// Mitsubishi GX Works2 project: plc_v1   PLC: Q03UDV

PROGRAM COM_RACK
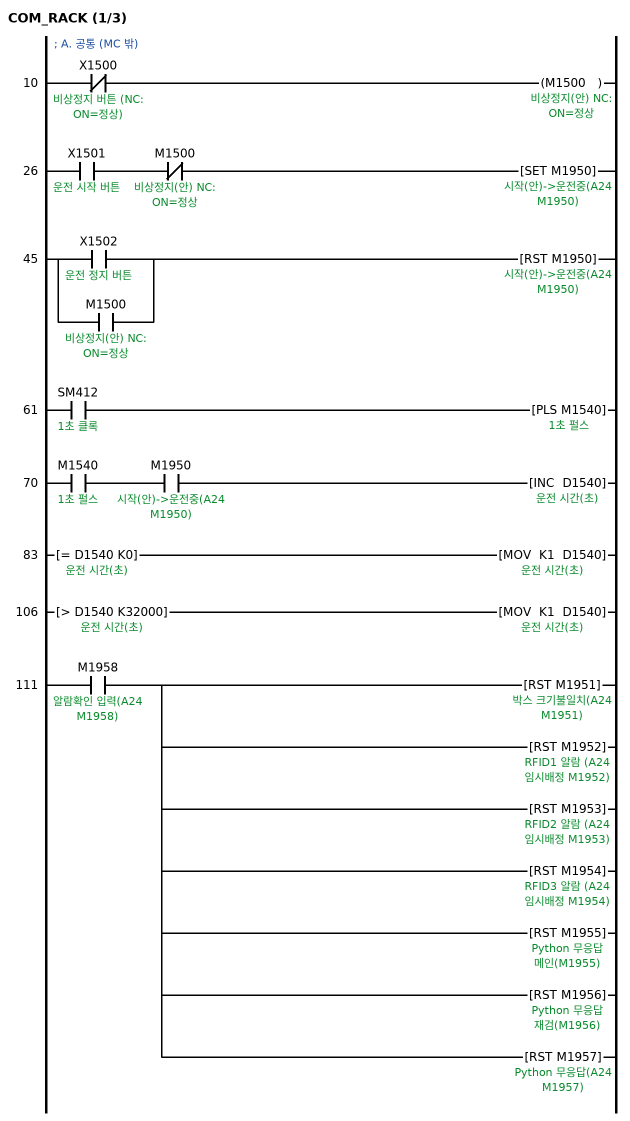
; A. 공통 (MC 밖)
10    LDI     X1500  ; 비상정지 버튼 (NC: ON=정상)
      OUT     M1500  ; 비상정지(안) NC: ON=정상
        [note] 비상정지(안) NC: ON=정상
26    LD      X1501  ; 운전 시작 버튼
      ANI     M1500  ; 비상정지(안) NC: ON=정상
      SET     M1950  ; 시작(안)->운전중(A24 M1950)
        [note] 시작(안)->운전중(A24 M1950)
45    LD      X1502  ; 운전 정지 버튼
      OR      M1500  ; 비상정지(안) NC: ON=정상
      RST     M1950  ; 시작(안)->운전중(A24 M1950)
        [note] 정지(안) 또는 비상정지
61    LD      SM412  ; 1초 클록
      PLS     M1540  ; 1초 펄스
        [note] 1초 펄스
70    LD      M1540  ; 1초 펄스
      AND     M1950  ; 시작(안)->운전중(A24 M1950)
      INC     D1540  ; 운전 시간(초)
        [note] 운전 시간(초)
83    LD=     D1540 K0  ; 운전 시간(초)
      MOV     K1 D1540
        [note] 0은 입고 중 표시로 쓰므로 1부터
106   LD>     D1540 K32000  ; 운전 시간(초)
      MOV     K1 D1540
111   LD      M1958  ; 알람확인 입력(A24 M1958)
      RST     M1951  ; 박스 크기불일치(A24 M1951)
      RST     M1952  ; RFID1 알람 (A24 임시배정 M1952)
      RST     M1953  ; RFID2 알람 (A24 임시배정 M1953)
      RST     M1954  ; RFID3 알람 (A24 임시배정 M1954)
      RST     M1955  ; Python 무응답 메인(M1955)
      RST     M1956  ; Python 무응답 재검(M1956)
      RST     M1957  ; Python 무응답(A24 M1957)
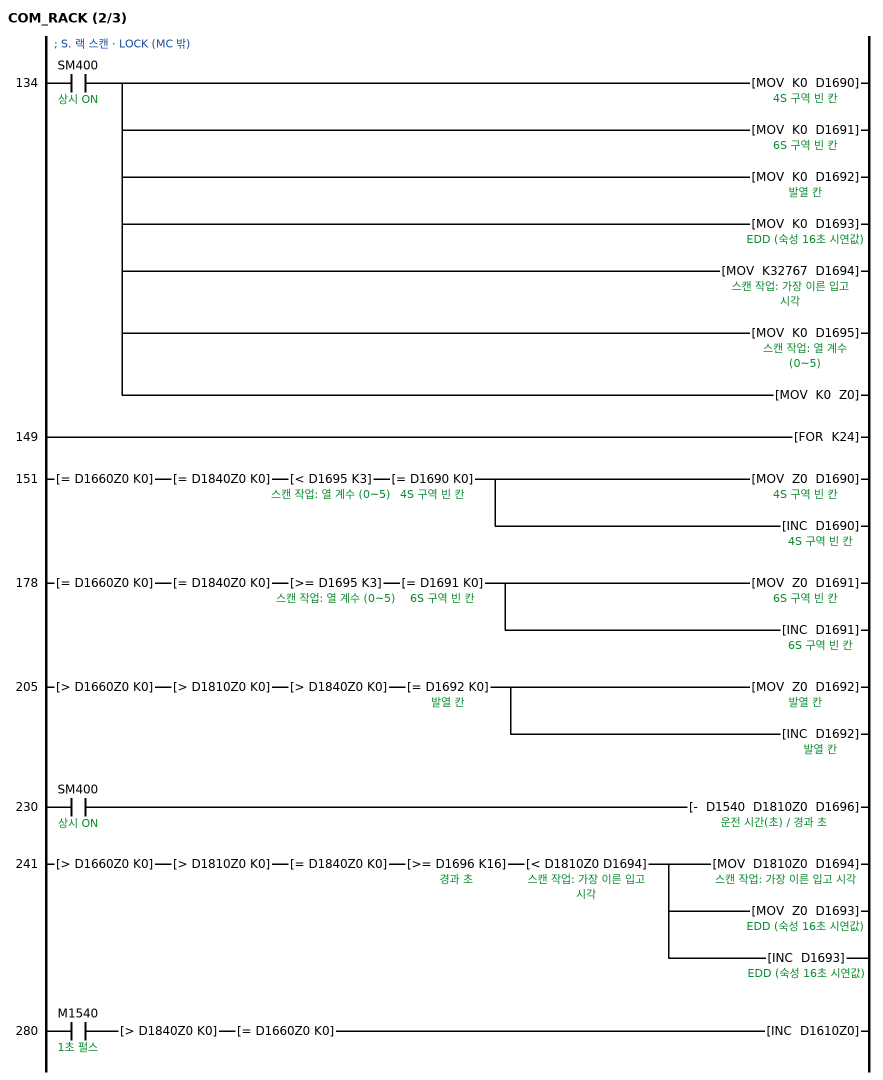
; S. 랙 스캔 · LOCK (MC 밖)
134   LD      SM400  ; 상시 ON
      MOV     K0 D1690  ; 4S 구역 빈 칸
      MOV     K0 D1691  ; 6S 구역 빈 칸
      MOV     K0 D1692  ; 발열 칸
      MOV     K0 D1693  ; EDD (숙성 16초 시연값)
      MOV     K32767 D1694  ; 스캔 작업: 가장 이른 입고 시각
      MOV     K0 D1695  ; 스캔 작업: 열 계수 (0~5)
      MOV     K0 Z0
149   FOR     K24
151   LD=     D1660Z0 K0
      AND=    D1840Z0 K0
      AND<    D1695 K3  ; 스캔 작업: 열 계수 (0~5)
      AND=    D1690 K0  ; 4S 구역 빈 칸
      MOV     Z0 D1690
      INC     D1690
        [note] 4S 구역 빈 칸
178   LD=     D1660Z0 K0
      AND=    D1840Z0 K0
      AND>=   D1695 K3  ; 스캔 작업: 열 계수 (0~5)
      AND=    D1691 K0  ; 6S 구역 빈 칸
      MOV     Z0 D1691
      INC     D1691
        [note] 6S 구역 빈 칸
205   LD>     D1660Z0 K0
      AND>    D1810Z0 K0
      AND>    D1840Z0 K0
      AND=    D1692 K0  ; 발열 칸
      MOV     Z0 D1692
      INC     D1692
        [note] 발열 칸
230   LD      SM400  ; 상시 ON
      -       D1540 D1810Z0 D1696  ; 경과 초
        [note] 경과 초
241   LD>     D1660Z0 K0
      AND>    D1810Z0 K0
      AND=    D1840Z0 K0
      AND>=   D1696 K16  ; 경과 초
      AND<    D1810Z0 D1694  ; 스캔 작업: 가장 이른 입고 시각
      MOV     D1810Z0 D1694
      MOV     Z0 D1693
      INC     D1693
        [note] EDD (숙성 16초 시연값)
280   LD      M1540  ; 1초 펄스
      AND>    D1840Z0 K0
      AND=    D1660Z0 K0
      INC     D1610Z0
        [note] LOCK 경과(초)
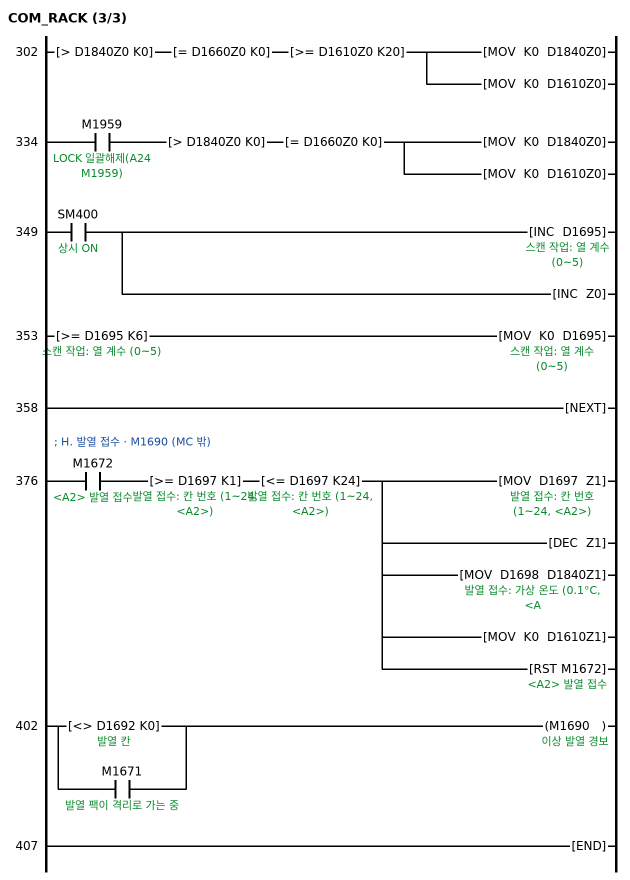
302   LD>     D1840Z0 K0
      AND=    D1660Z0 K0
      AND>=   D1610Z0 K20
      MOV     K0 D1840Z0
      MOV     K0 D1610Z0
        [note] 20초 뒤 자동 해제 (D13)
334   LD      M1959  ; LOCK 일괄해제(A24 M1959)
      AND>    D1840Z0 K0
      AND=    D1660Z0 K0
      MOV     K0 D1840Z0
      MOV     K0 D1610Z0
349   LD      SM400  ; 상시 ON
      INC     D1695
      INC     Z0
353   LD>=    D1695 K6  ; 스캔 작업: 열 계수 (0~5)
      MOV     K0 D1695
358   NEXT
; H. 발열 접수 · M1690 (MC 밖)
376   LD      M1672  ; <A2> 발열 접수
      AND>=   D1697 K1  ; 발열 접수: 칸 번호 (1~24, <A2>)
      AND<=   D1697 K24  ; 발열 접수: 칸 번호 (1~24, <A2>)
      MOV     D1697 Z1
      DEC     Z1
      MOV     D1698 D1840Z1  ; 발열 접수: 가상 온도 (0.1°C, <A
      MOV     K0 D1610Z1
      RST     M1672  ; <A2> 발열 접수
        [note] <A2> 발열 접수
402   LD<>    D1692 K0  ; 발열 칸
      OR      M1671  ; 발열 팩이 격리로 가는 중
      OUT     M1690  ; 이상 발열 경보
407   END
END_PROGRAM

PROGRAM MC_MAIN
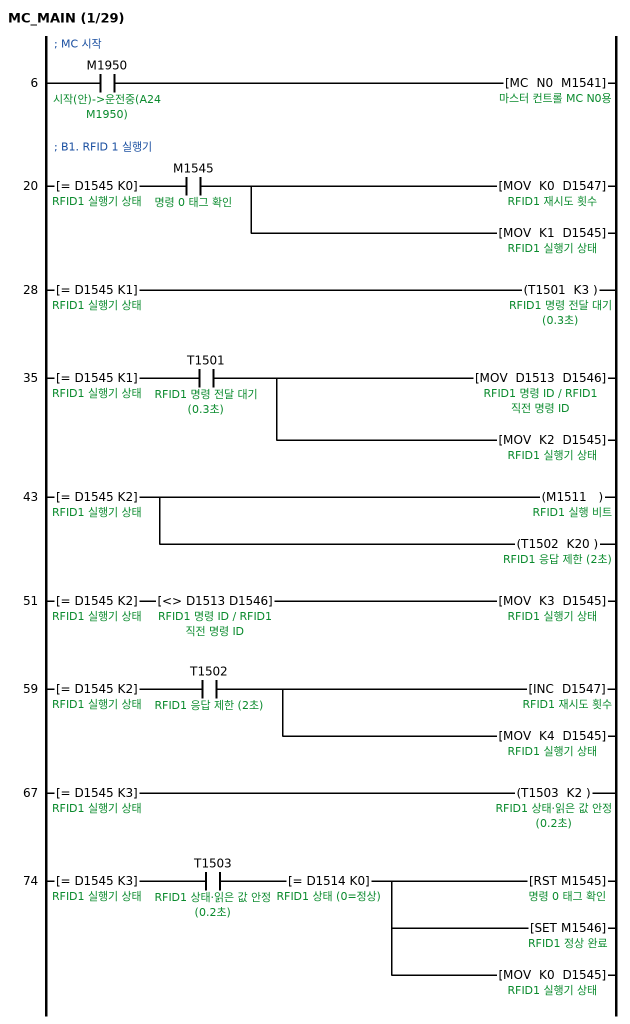
; MC 시작
6     LD      M1950  ; 시작(안)->운전중(A24 M1950)
      MC      N0 M1541  ; 마스터 컨트롤 MC N0용
; B1. RFID 1 실행기
20    LD=     D1545 K0  ; RFID1 실행기 상태
      AND     M1545  ; 명령 0 태그 확인
      MOV     K0 D1547  ; RFID1 재시도 횟수
      MOV     K1 D1545
28    LD=     D1545 K1  ; RFID1 실행기 상태
      OUT     T1501 K3  ; RFID1 명령 전달 대기 (0.3초)
35    LD=     D1545 K1  ; RFID1 실행기 상태
      AND     T1501  ; RFID1 명령 전달 대기 (0.3초)
      MOV     D1513 D1546  ; RFID1 명령 ID / RFID1 직전 명령 ID
      MOV     K2 D1545
43    LD=     D1545 K2  ; RFID1 실행기 상태
      OUT     M1511  ; RFID1 실행 비트
      OUT     T1502 K20  ; RFID1 응답 제한 (2초)
51    LD=     D1545 K2  ; RFID1 실행기 상태
      AND<>   D1513 D1546  ; RFID1 명령 ID / RFID1 직전 명령 ID
      MOV     K3 D1545
59    LD=     D1545 K2  ; RFID1 실행기 상태
      AND     T1502  ; RFID1 응답 제한 (2초)
      INC     D1547
      MOV     K4 D1545
67    LD=     D1545 K3  ; RFID1 실행기 상태
      OUT     T1503 K2  ; RFID1 상태·읽은 값 안정 (0.2초)
74    LD=     D1545 K3  ; RFID1 실행기 상태
      AND     T1503  ; RFID1 상태·읽은 값 안정 (0.2초)
      AND=    D1514 K0  ; RFID1 상태 (0=정상)
      RST     M1545  ; 명령 0 태그 확인
      SET     M1546  ; RFID1 정상 완료
      MOV     K0 D1545
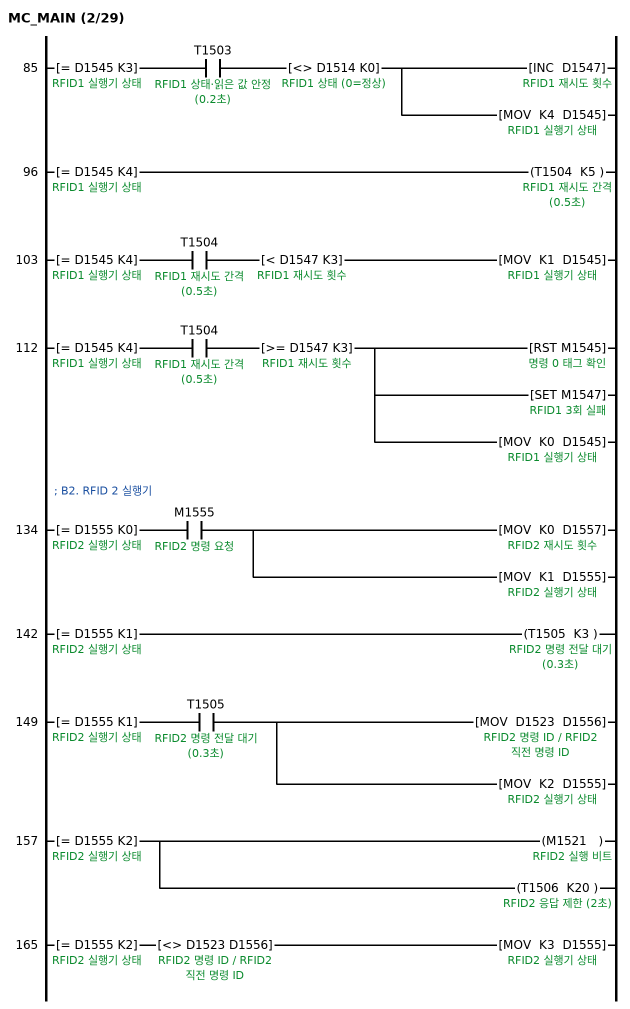
85    LD=     D1545 K3  ; RFID1 실행기 상태
      AND     T1503  ; RFID1 상태·읽은 값 안정 (0.2초)
      AND<>   D1514 K0  ; RFID1 상태 (0=정상)
      INC     D1547
      MOV     K4 D1545
96    LD=     D1545 K4  ; RFID1 실행기 상태
      OUT     T1504 K5  ; RFID1 재시도 간격 (0.5초)
103   LD=     D1545 K4  ; RFID1 실행기 상태
      AND     T1504  ; RFID1 재시도 간격 (0.5초)
      AND<    D1547 K3  ; RFID1 재시도 횟수
      MOV     K1 D1545
112   LD=     D1545 K4  ; RFID1 실행기 상태
      AND     T1504  ; RFID1 재시도 간격 (0.5초)
      AND>=   D1547 K3  ; RFID1 재시도 횟수
      RST     M1545  ; 명령 0 태그 확인
      SET     M1547  ; RFID1 3회 실패
      MOV     K0 D1545
; B2. RFID 2 실행기
134   LD=     D1555 K0  ; RFID2 실행기 상태
      AND     M1555  ; RFID2 명령 요청
      MOV     K0 D1557  ; RFID2 재시도 횟수
      MOV     K1 D1555
142   LD=     D1555 K1  ; RFID2 실행기 상태
      OUT     T1505 K3  ; RFID2 명령 전달 대기 (0.3초)
149   LD=     D1555 K1  ; RFID2 실행기 상태
      AND     T1505  ; RFID2 명령 전달 대기 (0.3초)
      MOV     D1523 D1556  ; RFID2 명령 ID / RFID2 직전 명령 ID
      MOV     K2 D1555
157   LD=     D1555 K2  ; RFID2 실행기 상태
      OUT     M1521  ; RFID2 실행 비트
      OUT     T1506 K20  ; RFID2 응답 제한 (2초)
165   LD=     D1555 K2  ; RFID2 실행기 상태
      AND<>   D1523 D1556  ; RFID2 명령 ID / RFID2 직전 명령 ID
      MOV     K3 D1555
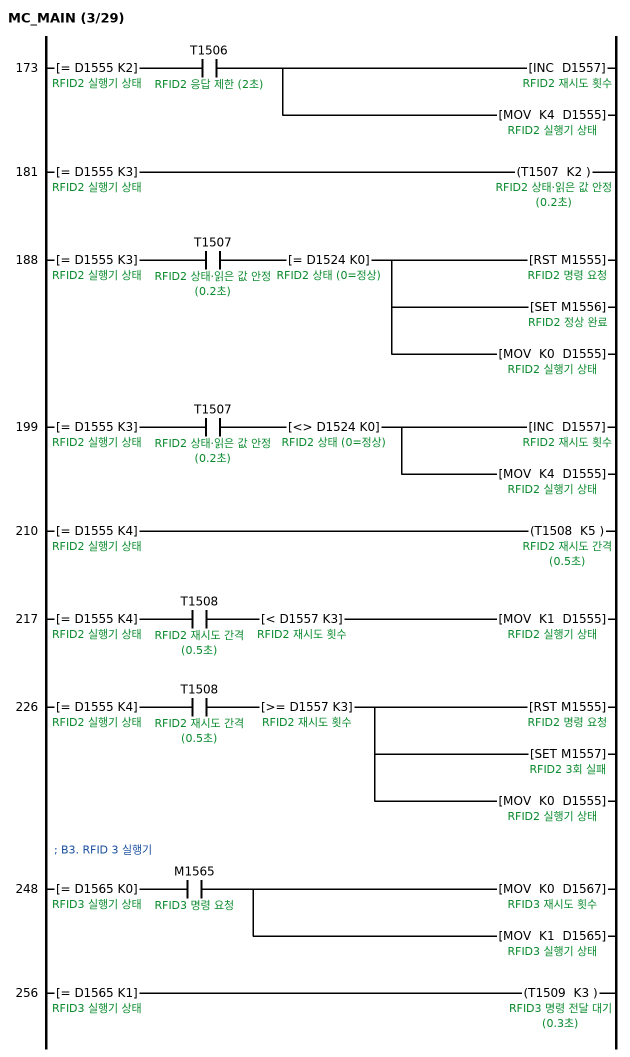
173   LD=     D1555 K2  ; RFID2 실행기 상태
      AND     T1506  ; RFID2 응답 제한 (2초)
      INC     D1557
      MOV     K4 D1555
181   LD=     D1555 K3  ; RFID2 실행기 상태
      OUT     T1507 K2  ; RFID2 상태·읽은 값 안정 (0.2초)
188   LD=     D1555 K3  ; RFID2 실행기 상태
      AND     T1507  ; RFID2 상태·읽은 값 안정 (0.2초)
      AND=    D1524 K0  ; RFID2 상태 (0=정상)
      RST     M1555  ; RFID2 명령 요청
      SET     M1556  ; RFID2 정상 완료
      MOV     K0 D1555
199   LD=     D1555 K3  ; RFID2 실행기 상태
      AND     T1507  ; RFID2 상태·읽은 값 안정 (0.2초)
      AND<>   D1524 K0  ; RFID2 상태 (0=정상)
      INC     D1557
      MOV     K4 D1555
210   LD=     D1555 K4  ; RFID2 실행기 상태
      OUT     T1508 K5  ; RFID2 재시도 간격 (0.5초)
217   LD=     D1555 K4  ; RFID2 실행기 상태
      AND     T1508  ; RFID2 재시도 간격 (0.5초)
      AND<    D1557 K3  ; RFID2 재시도 횟수
      MOV     K1 D1555
226   LD=     D1555 K4  ; RFID2 실행기 상태
      AND     T1508  ; RFID2 재시도 간격 (0.5초)
      AND>=   D1557 K3  ; RFID2 재시도 횟수
      RST     M1555  ; RFID2 명령 요청
      SET     M1557  ; RFID2 3회 실패
      MOV     K0 D1555
; B3. RFID 3 실행기
248   LD=     D1565 K0  ; RFID3 실행기 상태
      AND     M1565  ; RFID3 명령 요청
      MOV     K0 D1567  ; RFID3 재시도 횟수
      MOV     K1 D1565
256   LD=     D1565 K1  ; RFID3 실행기 상태
      OUT     T1509 K3  ; RFID3 명령 전달 대기 (0.3초)
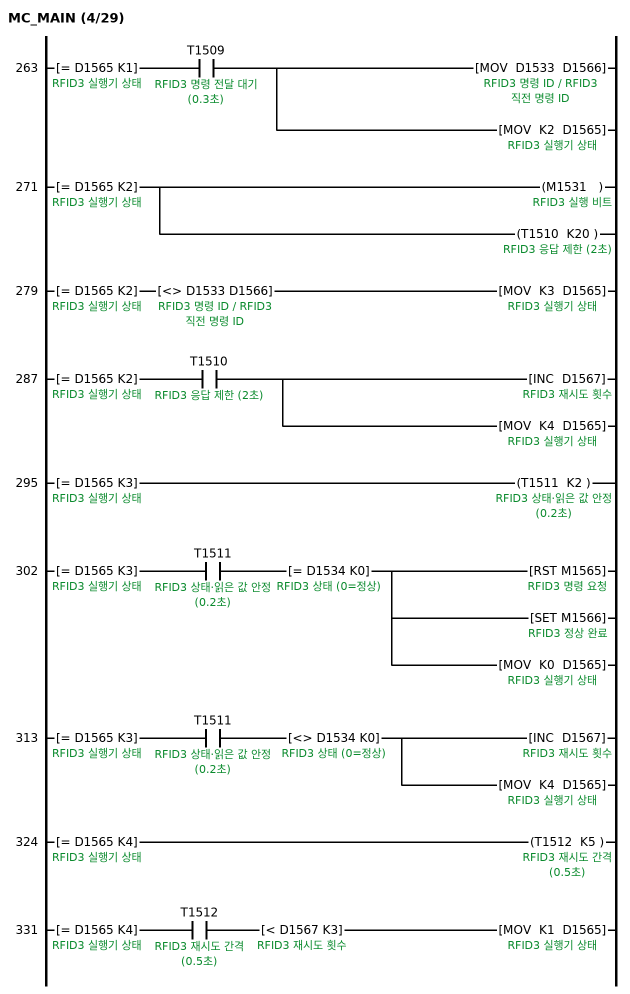
263   LD=     D1565 K1  ; RFID3 실행기 상태
      AND     T1509  ; RFID3 명령 전달 대기 (0.3초)
      MOV     D1533 D1566  ; RFID3 명령 ID / RFID3 직전 명령 ID
      MOV     K2 D1565
271   LD=     D1565 K2  ; RFID3 실행기 상태
      OUT     M1531  ; RFID3 실행 비트
      OUT     T1510 K20  ; RFID3 응답 제한 (2초)
279   LD=     D1565 K2  ; RFID3 실행기 상태
      AND<>   D1533 D1566  ; RFID3 명령 ID / RFID3 직전 명령 ID
      MOV     K3 D1565
287   LD=     D1565 K2  ; RFID3 실행기 상태
      AND     T1510  ; RFID3 응답 제한 (2초)
      INC     D1567
      MOV     K4 D1565
295   LD=     D1565 K3  ; RFID3 실행기 상태
      OUT     T1511 K2  ; RFID3 상태·읽은 값 안정 (0.2초)
302   LD=     D1565 K3  ; RFID3 실행기 상태
      AND     T1511  ; RFID3 상태·읽은 값 안정 (0.2초)
      AND=    D1534 K0  ; RFID3 상태 (0=정상)
      RST     M1565  ; RFID3 명령 요청
      SET     M1566  ; RFID3 정상 완료
      MOV     K0 D1565
313   LD=     D1565 K3  ; RFID3 실행기 상태
      AND     T1511  ; RFID3 상태·읽은 값 안정 (0.2초)
      AND<>   D1534 K0  ; RFID3 상태 (0=정상)
      INC     D1567
      MOV     K4 D1565
324   LD=     D1565 K4  ; RFID3 실행기 상태
      OUT     T1512 K5  ; RFID3 재시도 간격 (0.5초)
331   LD=     D1565 K4  ; RFID3 실행기 상태
      AND     T1512  ; RFID3 재시도 간격 (0.5초)
      AND<    D1567 K3  ; RFID3 재시도 횟수
      MOV     K1 D1565
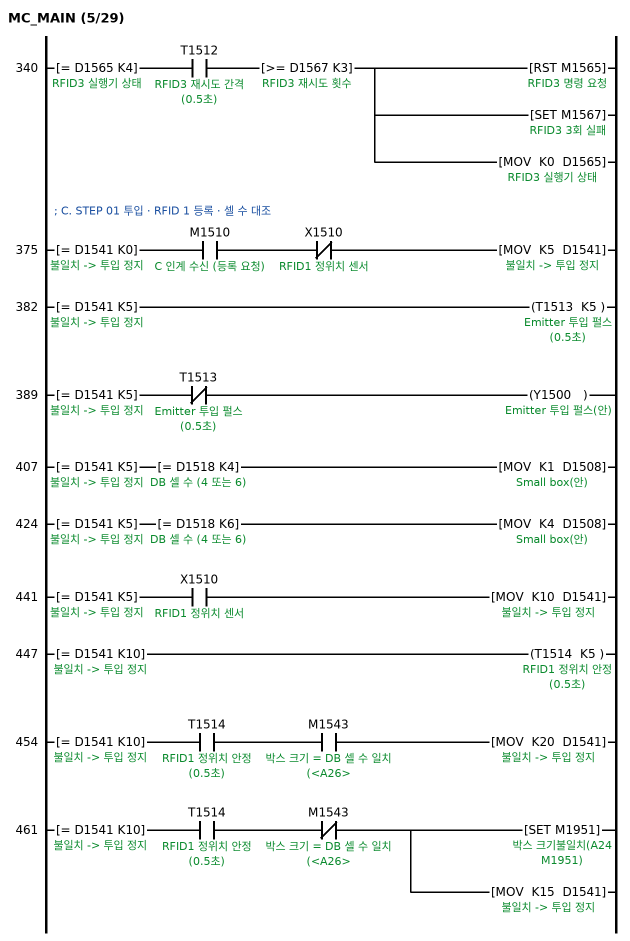
340   LD=     D1565 K4  ; RFID3 실행기 상태
      AND     T1512  ; RFID3 재시도 간격 (0.5초)
      AND>=   D1567 K3  ; RFID3 재시도 횟수
      RST     M1565  ; RFID3 명령 요청
      SET     M1567  ; RFID3 3회 실패
      MOV     K0 D1565
; C. STEP 01 투입 · RFID 1 등록 · 셀 수 대조
375   LD=     D1541 K0  ; 불일치 -> 투입 정지
      AND     M1510  ; C 인계 수신 (등록 요청)
      ANI     X1510  ; RFID1 정위치 센서
      MOV     K5 D1541
382   LD=     D1541 K5  ; 불일치 -> 투입 정지
      OUT     T1513 K5  ; Emitter 투입 펄스 (0.5초)
389   LD=     D1541 K5  ; 불일치 -> 투입 정지
      ANI     T1513  ; Emitter 투입 펄스 (0.5초)
      OUT     Y1500  ; Emitter 투입 펄스(안)
        [note] Emitter 투입 펄스(안)
407   LD=     D1541 K5  ; 불일치 -> 투입 정지
      AND=    D1518 K4  ; DB 셀 수 (4 또는 6)
      MOV     K1 D1508  ; Small box(안)
        [note] Small box(안)
424   LD=     D1541 K5  ; 불일치 -> 투입 정지
      AND=    D1518 K6  ; DB 셀 수 (4 또는 6)
      MOV     K4 D1508
        [note] Large box(안)
441   LD=     D1541 K5  ; 불일치 -> 투입 정지
      AND     X1510  ; RFID1 정위치 센서
      MOV     K10 D1541
447   LD=     D1541 K10  ; 불일치 -> 투입 정지
      OUT     T1514 K5  ; RFID1 정위치 안정 (0.5초)
454   LD=     D1541 K10  ; 불일치 -> 투입 정지
      AND     T1514  ; RFID1 정위치 안정 (0.5초)
      AND     M1543  ; 박스 크기 = DB 셀 수 일치 (<A26>
      MOV     K20 D1541
461   LD=     D1541 K10  ; 불일치 -> 투입 정지
      AND     T1514  ; RFID1 정위치 안정 (0.5초)
      ANI     M1543  ; 박스 크기 = DB 셀 수 일치 (<A26>
      SET     M1951  ; 박스 크기불일치(A24 M1951)
        [note] 박스 크기불일치(A24 M1951)
      MOV     K15 D1541
        [note] 불일치 -> 투입 정지
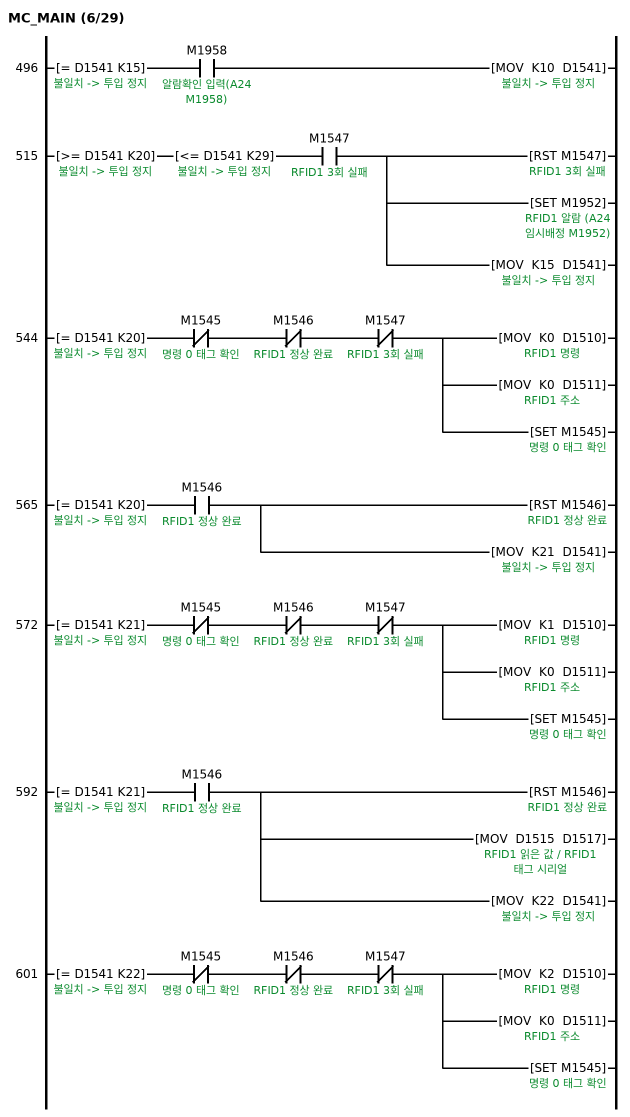
496   LD=     D1541 K15  ; 불일치 -> 투입 정지
      AND     M1958  ; 알람확인 입력(A24 M1958)
      MOV     K10 D1541
        [note] 알람 확인 뒤 다시 대조
515   LD>=    D1541 K20  ; 불일치 -> 투입 정지
      AND<=   D1541 K29  ; 불일치 -> 투입 정지
      AND     M1547  ; RFID1 3회 실패
      RST     M1547  ; RFID1 3회 실패
      SET     M1952  ; RFID1 알람 (A24 임시배정 M1952)
        [note] RFID1 알람 (A24 임시배정 M1952)
      MOV     K15 D1541
544   LD=     D1541 K20  ; 불일치 -> 투입 정지
      ANI     M1545  ; 명령 0 태그 확인
      ANI     M1546  ; RFID1 정상 완료
      ANI     M1547  ; RFID1 3회 실패
      MOV     K0 D1510  ; RFID1 명령
      MOV     K0 D1511  ; RFID1 주소
      SET     M1545  ; 명령 0 태그 확인
        [note] 명령 0 태그 확인
565   LD=     D1541 K20  ; 불일치 -> 투입 정지
      AND     M1546  ; RFID1 정상 완료
      RST     M1546  ; RFID1 정상 완료
      MOV     K21 D1541
572   LD=     D1541 K21  ; 불일치 -> 투입 정지
      ANI     M1545  ; 명령 0 태그 확인
      ANI     M1546  ; RFID1 정상 완료
      ANI     M1547  ; RFID1 3회 실패
      MOV     K1 D1510
      MOV     K0 D1511
      SET     M1545  ; 명령 0 태그 확인
        [note] 명령 1 시리얼
592   LD=     D1541 K21  ; 불일치 -> 투입 정지
      AND     M1546  ; RFID1 정상 완료
      RST     M1546  ; RFID1 정상 완료
      MOV     D1515 D1517  ; RFID1 읽은 값 / RFID1 태그 시리얼
      MOV     K22 D1541
601   LD=     D1541 K22  ; 불일치 -> 투입 정지
      ANI     M1545  ; 명령 0 태그 확인
      ANI     M1546  ; RFID1 정상 완료
      ANI     M1547  ; RFID1 3회 실패
      MOV     K2 D1510
      MOV     K0 D1511
      SET     M1545  ; 명령 0 태그 확인
        [note] 명령 2 idx0
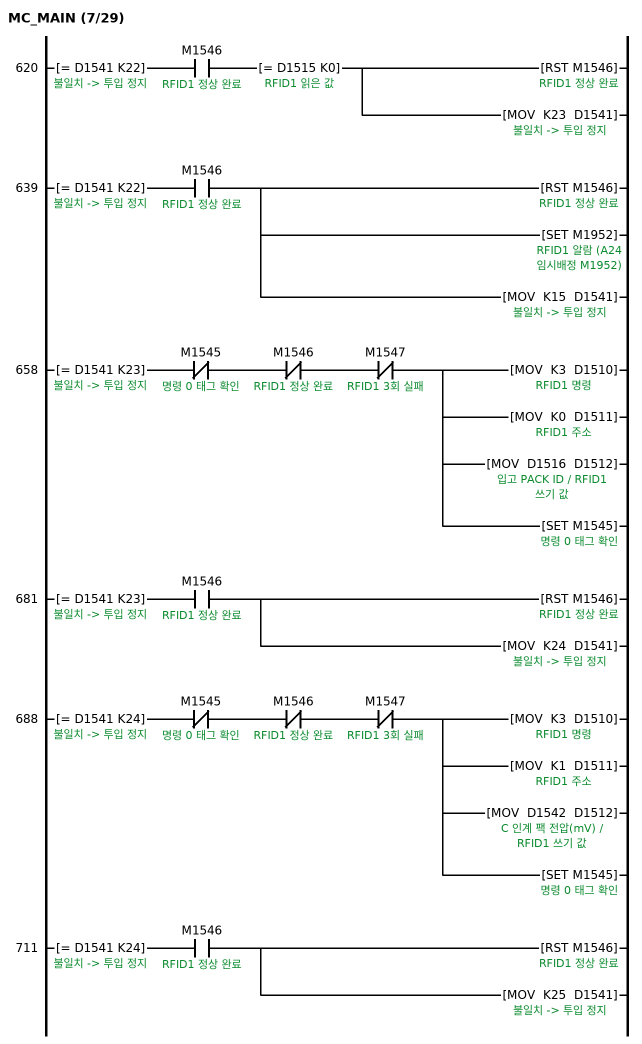
620   LD=     D1541 K22  ; 불일치 -> 투입 정지
      AND     M1546  ; RFID1 정상 완료
      AND=    D1515 K0  ; RFID1 읽은 값
      RST     M1546  ; RFID1 정상 완료
      MOV     K23 D1541
        [note] 미등록 -> 계속
639   LD=     D1541 K22  ; 불일치 -> 투입 정지
      AND     M1546  ; RFID1 정상 완료
      RST     M1546  ; RFID1 정상 완료
      SET     M1952  ; RFID1 알람 (A24 임시배정 M1952)
      MOV     K15 D1541
        [note] 0 아님 = 중복 투입
658   LD=     D1541 K23  ; 불일치 -> 투입 정지
      ANI     M1545  ; 명령 0 태그 확인
      ANI     M1546  ; RFID1 정상 완료
      ANI     M1547  ; RFID1 3회 실패
      MOV     K3 D1510
      MOV     K0 D1511
      MOV     D1516 D1512  ; 입고 PACK ID / RFID1 쓰기 값
      SET     M1545  ; 명령 0 태그 확인
        [note] idx0 <- PACK ID
681   LD=     D1541 K23  ; 불일치 -> 투입 정지
      AND     M1546  ; RFID1 정상 완료
      RST     M1546  ; RFID1 정상 완료
      MOV     K24 D1541
688   LD=     D1541 K24  ; 불일치 -> 투입 정지
      ANI     M1545  ; 명령 0 태그 확인
      ANI     M1546  ; RFID1 정상 완료
      ANI     M1547  ; RFID1 3회 실패
      MOV     K3 D1510
      MOV     K1 D1511
      MOV     D1542 D1512  ; C 인계 팩 전압(mV)
      SET     M1545  ; 명령 0 태그 확인
        [note] idx1 <- 팩 전압
711   LD=     D1541 K24  ; 불일치 -> 투입 정지
      AND     M1546  ; RFID1 정상 완료
      RST     M1546  ; RFID1 정상 완료
      MOV     K25 D1541
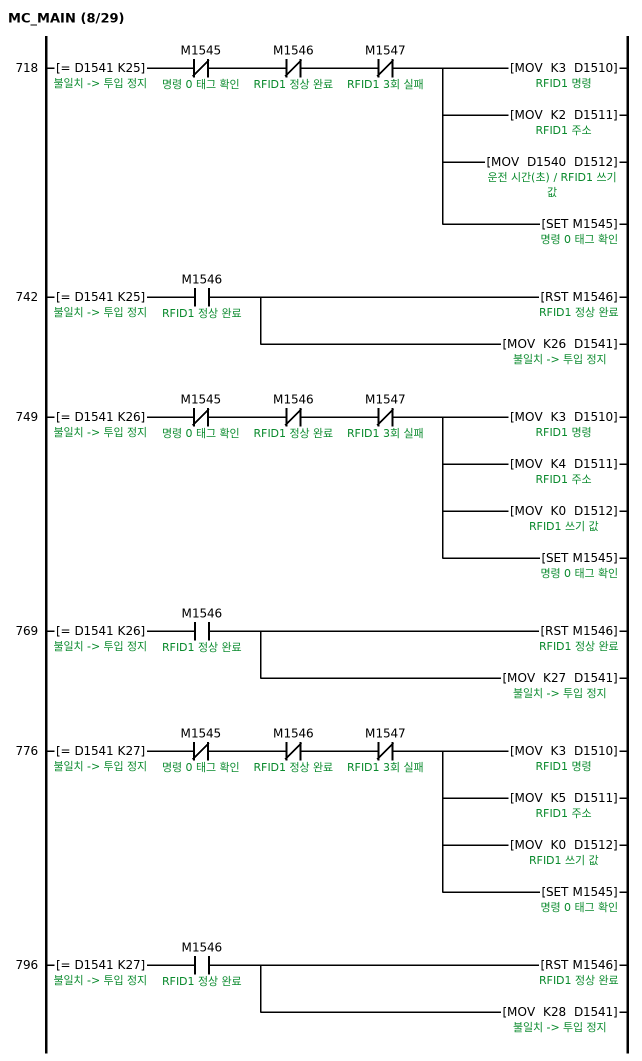
718   LD=     D1541 K25  ; 불일치 -> 투입 정지
      ANI     M1545  ; 명령 0 태그 확인
      ANI     M1546  ; RFID1 정상 완료
      ANI     M1547  ; RFID1 3회 실패
      MOV     K3 D1510
      MOV     K2 D1511
      MOV     D1540 D1512  ; 운전 시간(초)
      SET     M1545  ; 명령 0 태그 확인
        [note] idx2 <- 투입 시각
742   LD=     D1541 K25  ; 불일치 -> 투입 정지
      AND     M1546  ; RFID1 정상 완료
      RST     M1546  ; RFID1 정상 완료
      MOV     K26 D1541
749   LD=     D1541 K26  ; 불일치 -> 투입 정지
      ANI     M1545  ; 명령 0 태그 확인
      ANI     M1546  ; RFID1 정상 완료
      ANI     M1547  ; RFID1 3회 실패
      MOV     K3 D1510
      MOV     K4 D1511
      MOV     K0 D1512
      SET     M1545  ; 명령 0 태그 확인
        [note] idx4 <- 0
769   LD=     D1541 K26  ; 불일치 -> 투입 정지
      AND     M1546  ; RFID1 정상 완료
      RST     M1546  ; RFID1 정상 완료
      MOV     K27 D1541
776   LD=     D1541 K27  ; 불일치 -> 투입 정지
      ANI     M1545  ; 명령 0 태그 확인
      ANI     M1546  ; RFID1 정상 완료
      ANI     M1547  ; RFID1 3회 실패
      MOV     K3 D1510
      MOV     K5 D1511
      MOV     K0 D1512
      SET     M1545  ; 명령 0 태그 확인
        [note] idx5 <- 0
796   LD=     D1541 K27  ; 불일치 -> 투입 정지
      AND     M1546  ; RFID1 정상 완료
      RST     M1546  ; RFID1 정상 완료
      MOV     K28 D1541
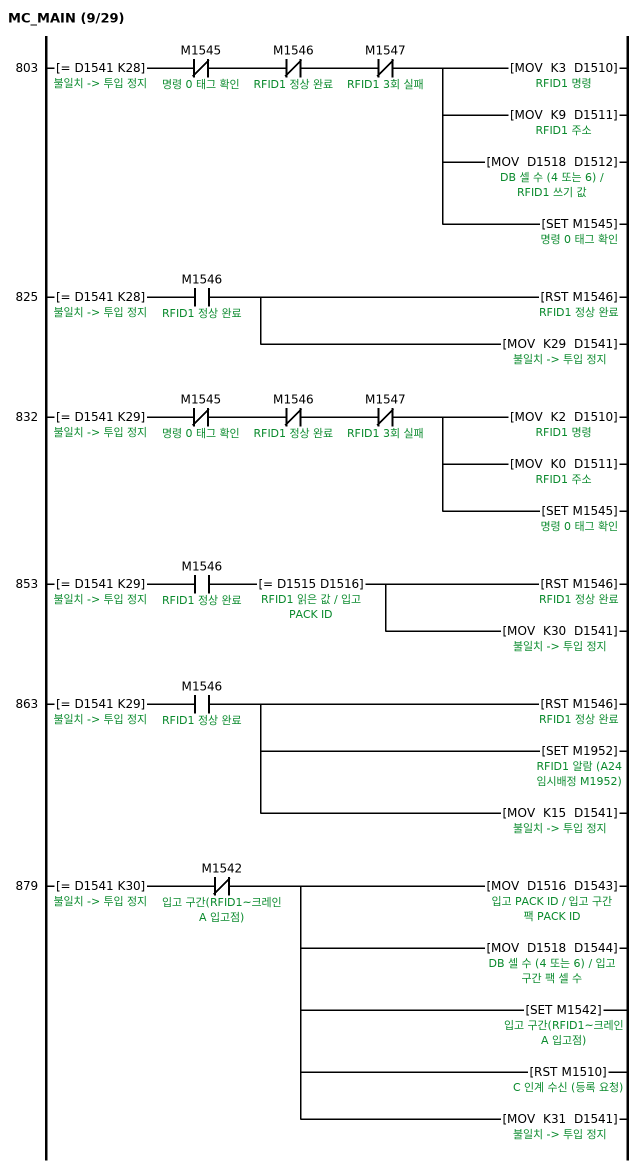
803   LD=     D1541 K28  ; 불일치 -> 투입 정지
      ANI     M1545  ; 명령 0 태그 확인
      ANI     M1546  ; RFID1 정상 완료
      ANI     M1547  ; RFID1 3회 실패
      MOV     K3 D1510
      MOV     K9 D1511
      MOV     D1518 D1512
      SET     M1545  ; 명령 0 태그 확인
        [note] idx9 <- 셀 수
825   LD=     D1541 K28  ; 불일치 -> 투입 정지
      AND     M1546  ; RFID1 정상 완료
      RST     M1546  ; RFID1 정상 완료
      MOV     K29 D1541
832   LD=     D1541 K29  ; 불일치 -> 투입 정지
      ANI     M1545  ; 명령 0 태그 확인
      ANI     M1546  ; RFID1 정상 완료
      ANI     M1547  ; RFID1 3회 실패
      MOV     K2 D1510
      MOV     K0 D1511
      SET     M1545  ; 명령 0 태그 확인
        [note] 명령 2 idx0 검증
853   LD=     D1541 K29  ; 불일치 -> 투입 정지
      AND     M1546  ; RFID1 정상 완료
      AND=    D1515 D1516  ; RFID1 읽은 값 / 입고 PACK ID
      RST     M1546  ; RFID1 정상 완료
      MOV     K30 D1541
863   LD=     D1541 K29  ; 불일치 -> 투입 정지
      AND     M1546  ; RFID1 정상 완료
      RST     M1546  ; RFID1 정상 완료
      SET     M1952  ; RFID1 알람 (A24 임시배정 M1952)
      MOV     K15 D1541
        [note] 검증 불일치
879   LD=     D1541 K30  ; 불일치 -> 투입 정지
      ANI     M1542  ; 입고 구간(RFID1~크레인A 입고점)
      MOV     D1516 D1543  ; 입고 구간 팩 PACK ID
      MOV     D1518 D1544  ; 입고 구간 팩 셀 수
      SET     M1542  ; 입고 구간(RFID1~크레인A 입고점)
      RST     M1510  ; C 인계 수신 (등록 요청)
      MOV     K31 D1541
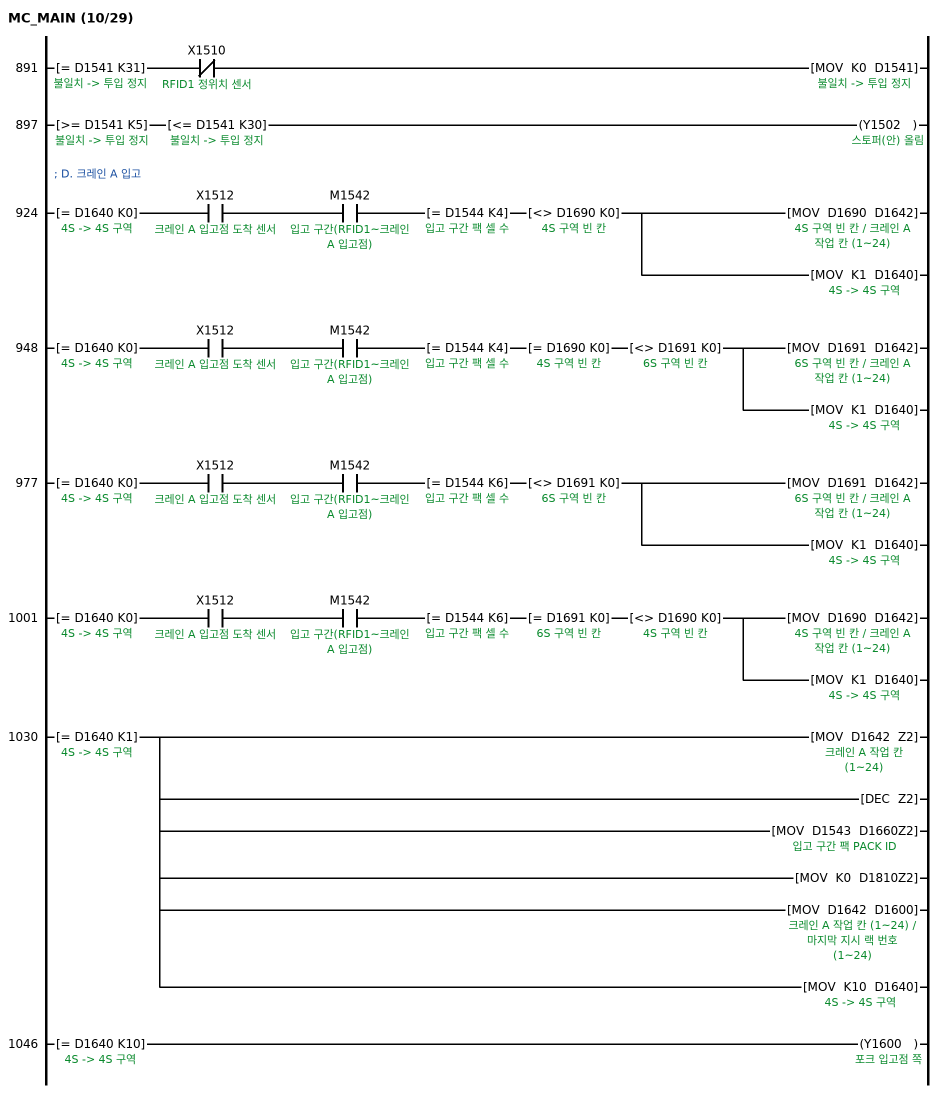
891   LD=     D1541 K31  ; 불일치 -> 투입 정지
      ANI     X1510  ; RFID1 정위치 센서
      MOV     K0 D1541
897   LD>=    D1541 K5  ; 불일치 -> 투입 정지
      AND<=   D1541 K30  ; 불일치 -> 투입 정지
      OUT     Y1502  ; 스토퍼(안) 올림
        [note] 스토퍼(안) 올림
; D. 크레인 A 입고
924   LD=     D1640 K0  ; 4S -> 4S 구역
      AND     X1512  ; 크레인 A 입고점 도착 센서
      AND     M1542  ; 입고 구간(RFID1~크레인A 입고점)
      AND=    D1544 K4  ; 입고 구간 팩 셀 수
      AND<>   D1690 K0  ; 4S 구역 빈 칸
      MOV     D1690 D1642  ; 크레인 A 작업 칸 (1~24)
      MOV     K1 D1640
        [note] 4S -> 4S 구역
948   LD=     D1640 K0  ; 4S -> 4S 구역
      AND     X1512  ; 크레인 A 입고점 도착 센서
      AND     M1542  ; 입고 구간(RFID1~크레인A 입고점)
      AND=    D1544 K4  ; 입고 구간 팩 셀 수
      AND=    D1690 K0  ; 4S 구역 빈 칸
      AND<>   D1691 K0  ; 6S 구역 빈 칸
      MOV     D1691 D1642
      MOV     K1 D1640
        [note] 4S 만차 -> 6S 구역
977   LD=     D1640 K0  ; 4S -> 4S 구역
      AND     X1512  ; 크레인 A 입고점 도착 센서
      AND     M1542  ; 입고 구간(RFID1~크레인A 입고점)
      AND=    D1544 K6  ; 입고 구간 팩 셀 수
      AND<>   D1691 K0  ; 6S 구역 빈 칸
      MOV     D1691 D1642
      MOV     K1 D1640
        [note] 6S -> 6S 구역
1001  LD=     D1640 K0  ; 4S -> 4S 구역
      AND     X1512  ; 크레인 A 입고점 도착 센서
      AND     M1542  ; 입고 구간(RFID1~크레인A 입고점)
      AND=    D1544 K6  ; 입고 구간 팩 셀 수
      AND=    D1691 K0  ; 6S 구역 빈 칸
      AND<>   D1690 K0  ; 4S 구역 빈 칸
      MOV     D1690 D1642
      MOV     K1 D1640
        [note] 6S 만차 -> 4S 구역
1030  LD=     D1640 K1  ; 4S -> 4S 구역
      MOV     D1642 Z2
      DEC     Z2
      MOV     D1543 D1660Z2
      MOV     K0 D1810Z2
      MOV     D1642 D1600  ; 마지막 지시 랙 번호 (1~24)
      MOV     K10 D1640
1046  LD=     D1640 K10  ; 4S -> 4S 구역
      OUT     Y1600  ; 포크 입고점 쪽
        [note] 포크 입고점 쪽
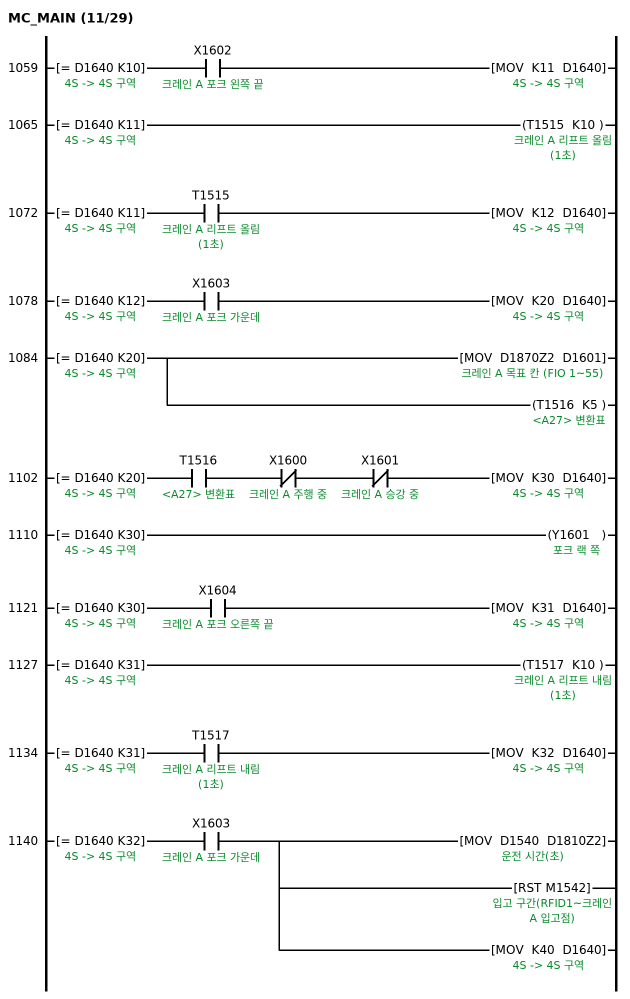
1059  LD=     D1640 K10  ; 4S -> 4S 구역
      AND     X1602  ; 크레인 A 포크 왼쪽 끝
      MOV     K11 D1640
1065  LD=     D1640 K11  ; 4S -> 4S 구역
      OUT     T1515 K10  ; 크레인 A 리프트 올림 (1초)
1072  LD=     D1640 K11  ; 4S -> 4S 구역
      AND     T1515  ; 크레인 A 리프트 올림 (1초)
      MOV     K12 D1640
1078  LD=     D1640 K12  ; 4S -> 4S 구역
      AND     X1603  ; 크레인 A 포크 가운데
      MOV     K20 D1640
1084  LD=     D1640 K20  ; 4S -> 4S 구역
      MOV     D1870Z2 D1601  ; 크레인 A 목표 칸 (FIO 1~55)
      OUT     T1516 K5  ; <A27> 변환표
        [note] <A27> 변환표
1102  LD=     D1640 K20  ; 4S -> 4S 구역
      AND     T1516  ; <A27> 변환표
      ANI     X1600  ; 크레인 A 주행 중
      ANI     X1601  ; 크레인 A 승강 중
      MOV     K30 D1640
1110  LD=     D1640 K30  ; 4S -> 4S 구역
      OUT     Y1601  ; 포크 랙 쪽
        [note] 포크 랙 쪽
1121  LD=     D1640 K30  ; 4S -> 4S 구역
      AND     X1604  ; 크레인 A 포크 오른쪽 끝
      MOV     K31 D1640
1127  LD=     D1640 K31  ; 4S -> 4S 구역
      OUT     T1517 K10  ; 크레인 A 리프트 내림 (1초)
1134  LD=     D1640 K31  ; 4S -> 4S 구역
      AND     T1517  ; 크레인 A 리프트 내림 (1초)
      MOV     K32 D1640
1140  LD=     D1640 K32  ; 4S -> 4S 구역
      AND     X1603  ; 크레인 A 포크 가운데
      MOV     D1540 D1810Z2
      RST     M1542  ; 입고 구간(RFID1~크레인A 입고점)
      MOV     K40 D1640
        [note] 입고 시각 = 숙성 시작
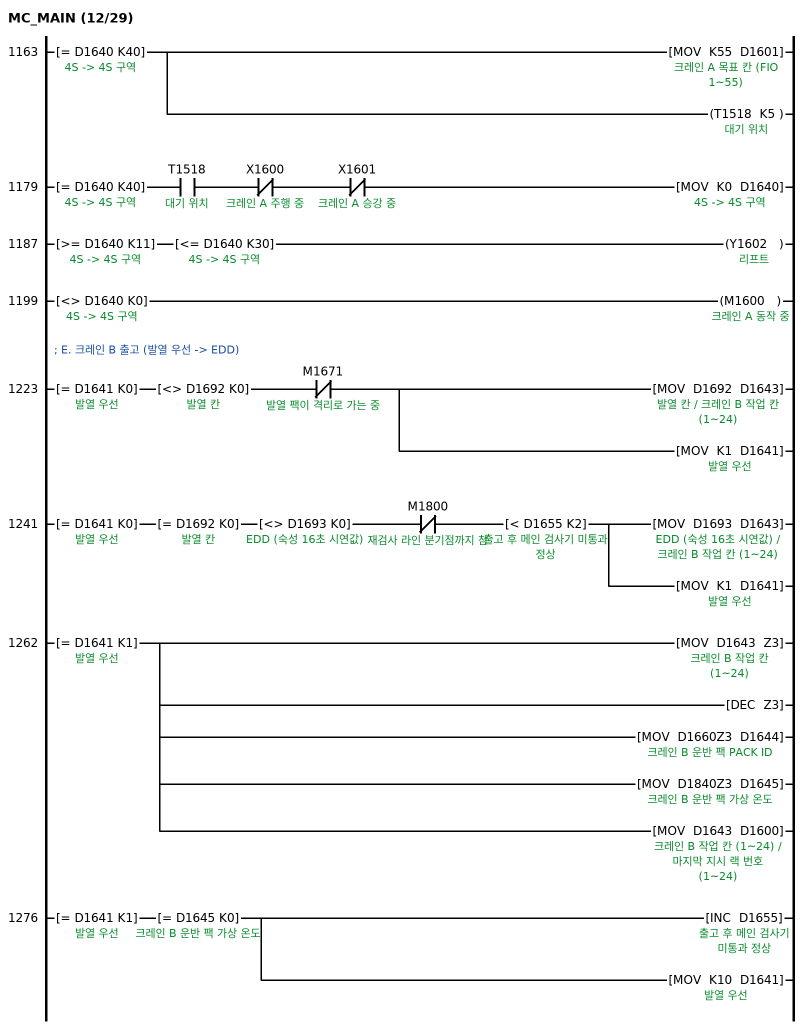
1163  LD=     D1640 K40  ; 4S -> 4S 구역
      MOV     K55 D1601
      OUT     T1518 K5  ; 대기 위치
        [note] 대기 위치
1179  LD=     D1640 K40  ; 4S -> 4S 구역
      AND     T1518  ; 대기 위치
      ANI     X1600  ; 크레인 A 주행 중
      ANI     X1601  ; 크레인 A 승강 중
      MOV     K0 D1640
1187  LD>=    D1640 K11  ; 4S -> 4S 구역
      AND<=   D1640 K30  ; 4S -> 4S 구역
      OUT     Y1602  ; 리프트
        [note] 리프트
1199  LD<>    D1640 K0  ; 4S -> 4S 구역
      OUT     M1600  ; 크레인 A 동작 중
; E. 크레인 B 출고 (발열 우선 -> EDD)
1223  LD=     D1641 K0  ; 발열 우선
      AND<>   D1692 K0  ; 발열 칸
      ANI     M1671  ; 발열 팩이 격리로 가는 중
      MOV     D1692 D1643  ; 크레인 B 작업 칸 (1~24)
      MOV     K1 D1641
        [note] 발열 우선
1241  LD=     D1641 K0  ; 발열 우선
      AND=    D1692 K0  ; 발열 칸
      AND<>   D1693 K0  ; EDD (숙성 16초 시연값)
      ANI     M1800  ; 재검사 라인 분기점까지 참
      AND<    D1655 K2  ; 출고 후 메인 검사기 미통과 정상
      MOV     D1693 D1643
      MOV     K1 D1641
        [note] EDD
1262  LD=     D1641 K1  ; 발열 우선
      MOV     D1643 Z3
      DEC     Z3
      MOV     D1660Z3 D1644  ; 크레인 B 운반 팩 PACK ID
      MOV     D1840Z3 D1645  ; 크레인 B 운반 팩 가상 온도
      MOV     D1643 D1600
1276  LD=     D1641 K1  ; 발열 우선
      AND=    D1645 K0  ; 크레인 B 운반 팩 가상 온도
      INC     D1655
      MOV     K10 D1641
        [note] 정상 팩
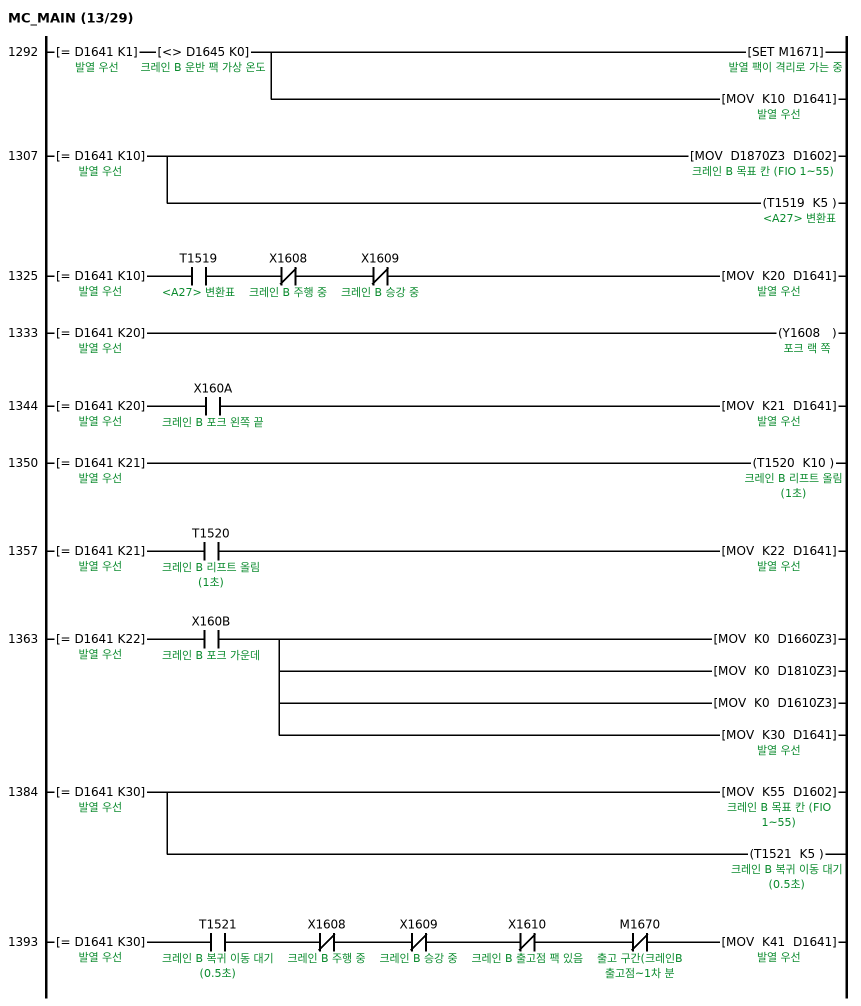
1292  LD=     D1641 K1  ; 발열 우선
      AND<>   D1645 K0  ; 크레인 B 운반 팩 가상 온도
      SET     M1671  ; 발열 팩이 격리로 가는 중
      MOV     K10 D1641
        [note] 발열 팩
1307  LD=     D1641 K10  ; 발열 우선
      MOV     D1870Z3 D1602  ; 크레인 B 목표 칸 (FIO 1~55)
      OUT     T1519 K5  ; <A27> 변환표
        [note] <A27> 변환표
1325  LD=     D1641 K10  ; 발열 우선
      AND     T1519  ; <A27> 변환표
      ANI     X1608  ; 크레인 B 주행 중
      ANI     X1609  ; 크레인 B 승강 중
      MOV     K20 D1641
1333  LD=     D1641 K20  ; 발열 우선
      OUT     Y1608  ; 포크 랙 쪽
        [note] 포크 랙 쪽
1344  LD=     D1641 K20  ; 발열 우선
      AND     X160A  ; 크레인 B 포크 왼쪽 끝
      MOV     K21 D1641
1350  LD=     D1641 K21  ; 발열 우선
      OUT     T1520 K10  ; 크레인 B 리프트 올림 (1초)
1357  LD=     D1641 K21  ; 발열 우선
      AND     T1520  ; 크레인 B 리프트 올림 (1초)
      MOV     K22 D1641
1363  LD=     D1641 K22  ; 발열 우선
      AND     X160B  ; 크레인 B 포크 가운데
      MOV     K0 D1660Z3
      MOV     K0 D1810Z3
      MOV     K0 D1610Z3
      MOV     K30 D1641
        [note] 칸 비움
1384  LD=     D1641 K30  ; 발열 우선
      MOV     K55 D1602
      OUT     T1521 K5  ; 크레인 B 복귀 이동 대기 (0.5초)
1393  LD=     D1641 K30  ; 발열 우선
      AND     T1521  ; 크레인 B 복귀 이동 대기 (0.5초)
      ANI     X1608  ; 크레인 B 주행 중
      ANI     X1609  ; 크레인 B 승강 중
      ANI     X1610  ; 크레인 B 출고점 팩 있음
      ANI     M1670  ; 출고 구간(크레인B 출고점~1차 분
      MOV     K41 D1641
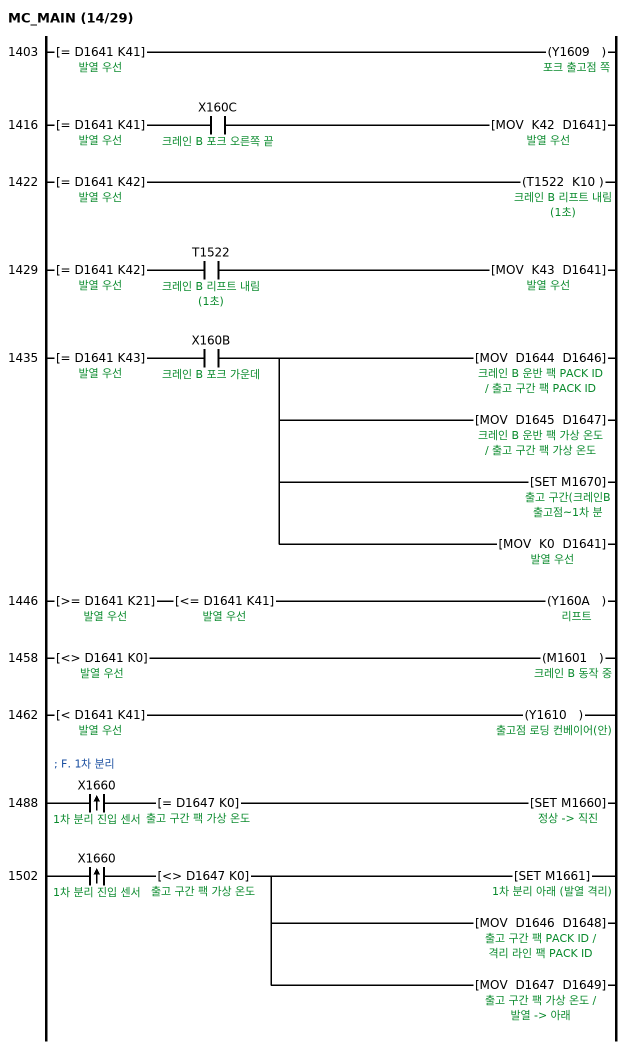
1403  LD=     D1641 K41  ; 발열 우선
      OUT     Y1609  ; 포크 출고점 쪽
        [note] 포크 출고점 쪽
1416  LD=     D1641 K41  ; 발열 우선
      AND     X160C  ; 크레인 B 포크 오른쪽 끝
      MOV     K42 D1641
1422  LD=     D1641 K42  ; 발열 우선
      OUT     T1522 K10  ; 크레인 B 리프트 내림 (1초)
1429  LD=     D1641 K42  ; 발열 우선
      AND     T1522  ; 크레인 B 리프트 내림 (1초)
      MOV     K43 D1641
1435  LD=     D1641 K43  ; 발열 우선
      AND     X160B  ; 크레인 B 포크 가운데
      MOV     D1644 D1646  ; 출고 구간 팩 PACK ID
      MOV     D1645 D1647  ; 출고 구간 팩 가상 온도
      SET     M1670  ; 출고 구간(크레인B 출고점~1차 분
      MOV     K0 D1641
1446  LD>=    D1641 K21  ; 발열 우선
      AND<=   D1641 K41  ; 발열 우선
      OUT     Y160A  ; 리프트
        [note] 리프트
1458  LD<>    D1641 K0  ; 발열 우선
      OUT     M1601  ; 크레인 B 동작 중
1462  LD<     D1641 K41  ; 발열 우선
      OUT     Y1610  ; 출고점 로딩 컨베이어(안)
        [note] 출고점 로딩 컨베이어(안)
; F. 1차 분리
1488  LDP     X1660  ; 1차 분리 진입 센서
      AND=    D1647 K0  ; 출고 구간 팩 가상 온도
      SET     M1660  ; 정상 -> 직진
        [note] 정상 -> 직진
1502  LDP     X1660  ; 1차 분리 진입 센서
      AND<>   D1647 K0  ; 출고 구간 팩 가상 온도
      SET     M1661  ; 1차 분리 아래 (발열 격리)
      MOV     D1646 D1648  ; 격리 라인 팩 PACK ID
      MOV     D1647 D1649  ; 발열 -> 아래
        [note] 발열 -> 아래
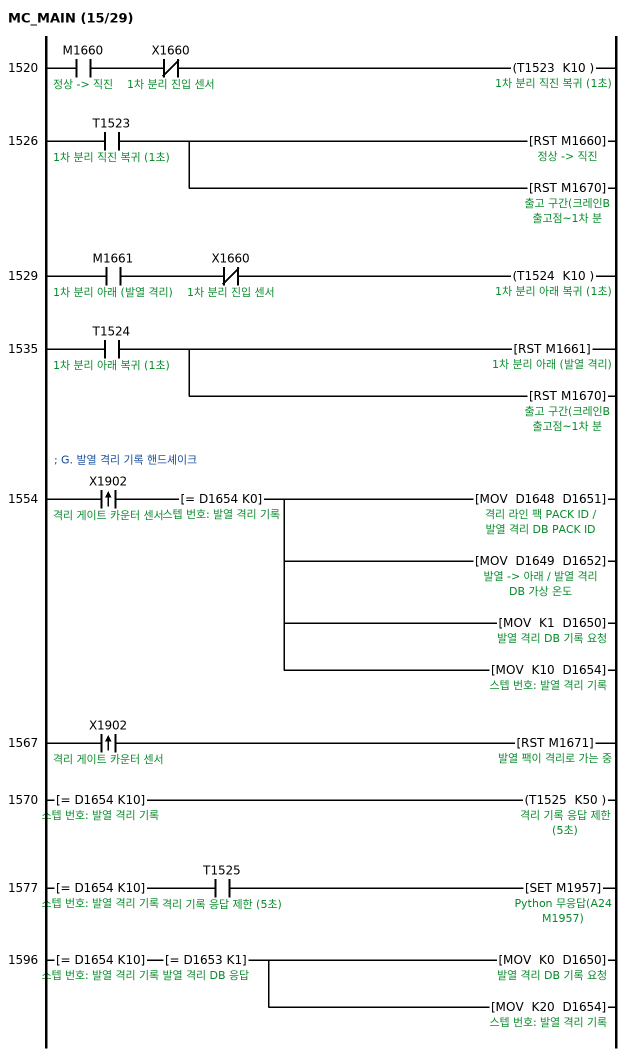
1520  LD      M1660  ; 정상 -> 직진
      ANI     X1660  ; 1차 분리 진입 센서
      OUT     T1523 K10  ; 1차 분리 직진 복귀 (1초)
1526  LD      T1523  ; 1차 분리 직진 복귀 (1초)
      RST     M1660  ; 정상 -> 직진
      RST     M1670  ; 출고 구간(크레인B 출고점~1차 분
1529  LD      M1661  ; 1차 분리 아래 (발열 격리)
      ANI     X1660  ; 1차 분리 진입 센서
      OUT     T1524 K10  ; 1차 분리 아래 복귀 (1초)
1535  LD      T1524  ; 1차 분리 아래 복귀 (1초)
      RST     M1661  ; 1차 분리 아래 (발열 격리)
      RST     M1670  ; 출고 구간(크레인B 출고점~1차 분
; G. 발열 격리 기록 핸드셰이크
1554  LDP     X1902  ; 격리 게이트 카운터 센서
      AND=    D1654 K0  ; 스텝 번호: 발열 격리 기록
      MOV     D1648 D1651  ; 발열 격리 DB PACK ID
      MOV     D1649 D1652  ; 발열 격리 DB 가상 온도
      MOV     K1 D1650  ; 발열 격리 DB 기록 요청
      MOV     K10 D1654
1567  LDP     X1902  ; 격리 게이트 카운터 센서
      RST     M1671  ; 발열 팩이 격리로 가는 중
1570  LD=     D1654 K10  ; 스텝 번호: 발열 격리 기록
      OUT     T1525 K50  ; 격리 기록 응답 제한 (5초)
1577  LD=     D1654 K10  ; 스텝 번호: 발열 격리 기록
      AND     T1525  ; 격리 기록 응답 제한 (5초)
      SET     M1957  ; Python 무응답(A24 M1957)
        [note] Python 무응답(A24 M1957)
1596  LD=     D1654 K10  ; 스텝 번호: 발열 격리 기록
      AND=    D1653 K1  ; 발열 격리 DB 응답
      MOV     K0 D1650
      MOV     K20 D1654
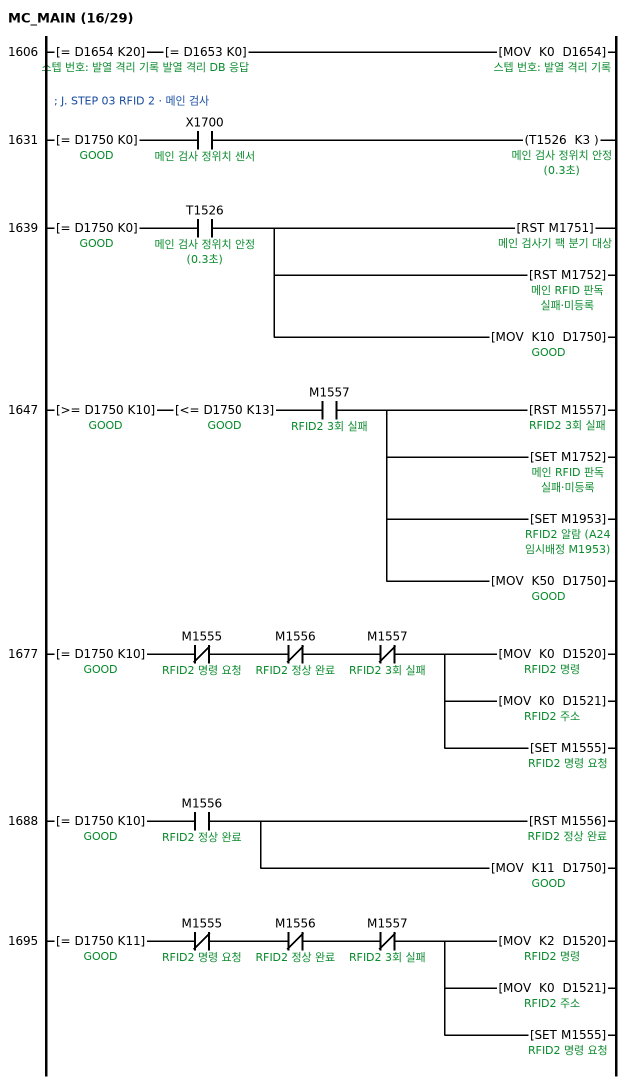
1606  LD=     D1654 K20  ; 스텝 번호: 발열 격리 기록
      AND=    D1653 K0  ; 발열 격리 DB 응답
      MOV     K0 D1654
; J. STEP 03 RFID 2 · 메인 검사
1631  LD=     D1750 K0  ; GOOD
      AND     X1700  ; 메인 검사 정위치 센서
      OUT     T1526 K3  ; 메인 검사 정위치 안정 (0.3초)
1639  LD=     D1750 K0  ; GOOD
      AND     T1526  ; 메인 검사 정위치 안정 (0.3초)
      RST     M1751  ; 메인 검사기 팩 분기 대상
      RST     M1752  ; 메인 RFID 판독 실패·미등록
      MOV     K10 D1750
1647  LD>=    D1750 K10  ; GOOD
      AND<=   D1750 K13  ; GOOD
      AND     M1557  ; RFID2 3회 실패
      RST     M1557  ; RFID2 3회 실패
      SET     M1752  ; 메인 RFID 판독 실패·미등록
      SET     M1953  ; RFID2 알람 (A24 임시배정 M1953)
        [note] RFID2 알람 (A24 임시배정 M1953)
      MOV     K50 D1750
1677  LD=     D1750 K10  ; GOOD
      ANI     M1555  ; RFID2 명령 요청
      ANI     M1556  ; RFID2 정상 완료
      ANI     M1557  ; RFID2 3회 실패
      MOV     K0 D1520  ; RFID2 명령
      MOV     K0 D1521  ; RFID2 주소
      SET     M1555  ; RFID2 명령 요청
1688  LD=     D1750 K10  ; GOOD
      AND     M1556  ; RFID2 정상 완료
      RST     M1556  ; RFID2 정상 완료
      MOV     K11 D1750
1695  LD=     D1750 K11  ; GOOD
      ANI     M1555  ; RFID2 명령 요청
      ANI     M1556  ; RFID2 정상 완료
      ANI     M1557  ; RFID2 3회 실패
      MOV     K2 D1520
      MOV     K0 D1521
      SET     M1555  ; RFID2 명령 요청
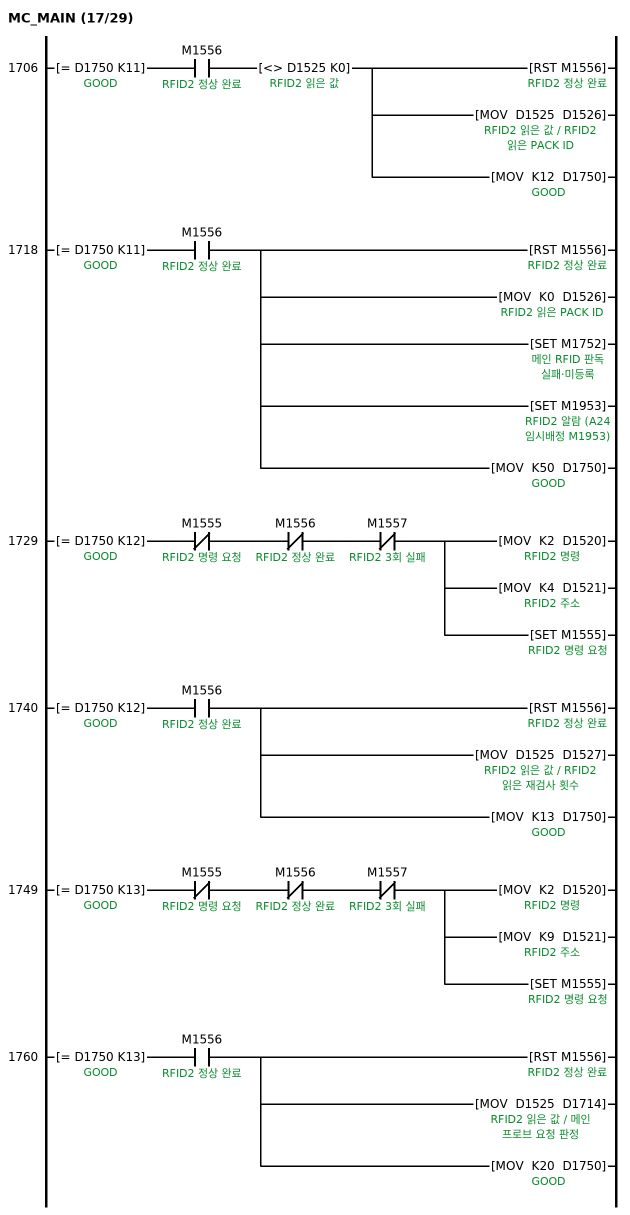
1706  LD=     D1750 K11  ; GOOD
      AND     M1556  ; RFID2 정상 완료
      AND<>   D1525 K0  ; RFID2 읽은 값
      RST     M1556  ; RFID2 정상 완료
      MOV     D1525 D1526  ; RFID2 읽은 PACK ID
      MOV     K12 D1750
1718  LD=     D1750 K11  ; GOOD
      AND     M1556  ; RFID2 정상 완료
      RST     M1556  ; RFID2 정상 완료
      MOV     K0 D1526
      SET     M1752  ; 메인 RFID 판독 실패·미등록
      SET     M1953  ; RFID2 알람 (A24 임시배정 M1953)
      MOV     K50 D1750
1729  LD=     D1750 K12  ; GOOD
      ANI     M1555  ; RFID2 명령 요청
      ANI     M1556  ; RFID2 정상 완료
      ANI     M1557  ; RFID2 3회 실패
      MOV     K2 D1520
      MOV     K4 D1521
      SET     M1555  ; RFID2 명령 요청
1740  LD=     D1750 K12  ; GOOD
      AND     M1556  ; RFID2 정상 완료
      RST     M1556  ; RFID2 정상 완료
      MOV     D1525 D1527  ; RFID2 읽은 재검사 횟수
      MOV     K13 D1750
1749  LD=     D1750 K13  ; GOOD
      ANI     M1555  ; RFID2 명령 요청
      ANI     M1556  ; RFID2 정상 완료
      ANI     M1557  ; RFID2 3회 실패
      MOV     K2 D1520
      MOV     K9 D1521
      SET     M1555  ; RFID2 명령 요청
1760  LD=     D1750 K13  ; GOOD
      AND     M1556  ; RFID2 정상 완료
      RST     M1556  ; RFID2 정상 완료
      MOV     D1525 D1714  ; 메인 프로브 요청 판정
      MOV     K20 D1750
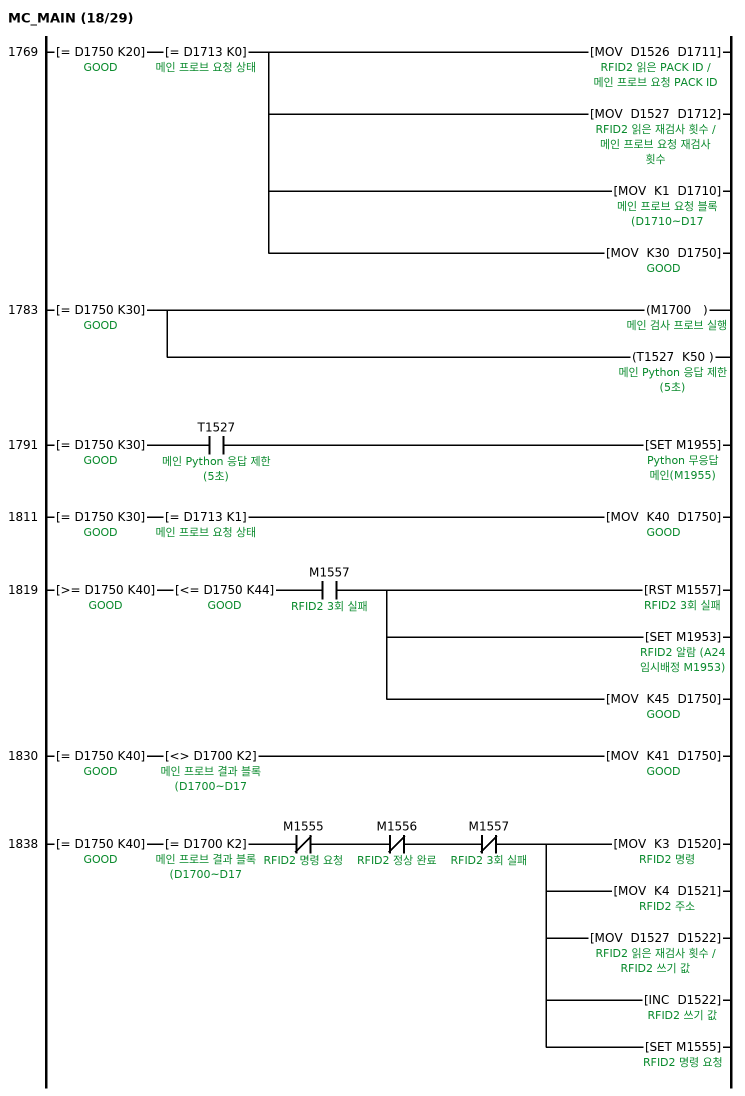
1769  LD=     D1750 K20  ; GOOD
      AND=    D1713 K0  ; 메인 프로브 요청 상태
      MOV     D1526 D1711  ; 메인 프로브 요청 PACK ID
      MOV     D1527 D1712  ; 메인 프로브 요청 재검사 횟수
      MOV     K1 D1710  ; 메인 프로브 요청 블록 (D1710~D17
      MOV     K30 D1750
1783  LD=     D1750 K30  ; GOOD
      OUT     M1700  ; 메인 검사 프로브 실행
      OUT     T1527 K50  ; 메인 Python 응답 제한 (5초)
1791  LD=     D1750 K30  ; GOOD
      AND     T1527  ; 메인 Python 응답 제한 (5초)
      SET     M1955  ; Python 무응답 메인(M1955)
        [note] Python 무응답 메인(M1955)
1811  LD=     D1750 K30  ; GOOD
      AND=    D1713 K1  ; 메인 프로브 요청 상태
      MOV     K40 D1750
1819  LD>=    D1750 K40  ; GOOD
      AND<=   D1750 K44  ; GOOD
      AND     M1557  ; RFID2 3회 실패
      RST     M1557  ; RFID2 3회 실패
      SET     M1953  ; RFID2 알람 (A24 임시배정 M1953)
      MOV     K45 D1750
1830  LD=     D1750 K40  ; GOOD
      AND<>   D1700 K2  ; 메인 프로브 결과 블록 (D1700~D17
      MOV     K41 D1750
1838  LD=     D1750 K40  ; GOOD
      AND=    D1700 K2  ; 메인 프로브 결과 블록 (D1700~D17
      ANI     M1555  ; RFID2 명령 요청
      ANI     M1556  ; RFID2 정상 완료
      ANI     M1557  ; RFID2 3회 실패
      MOV     K3 D1520
      MOV     K4 D1521
      MOV     D1527 D1522  ; RFID2 쓰기 값
      INC     D1522
      SET     M1555  ; RFID2 명령 요청
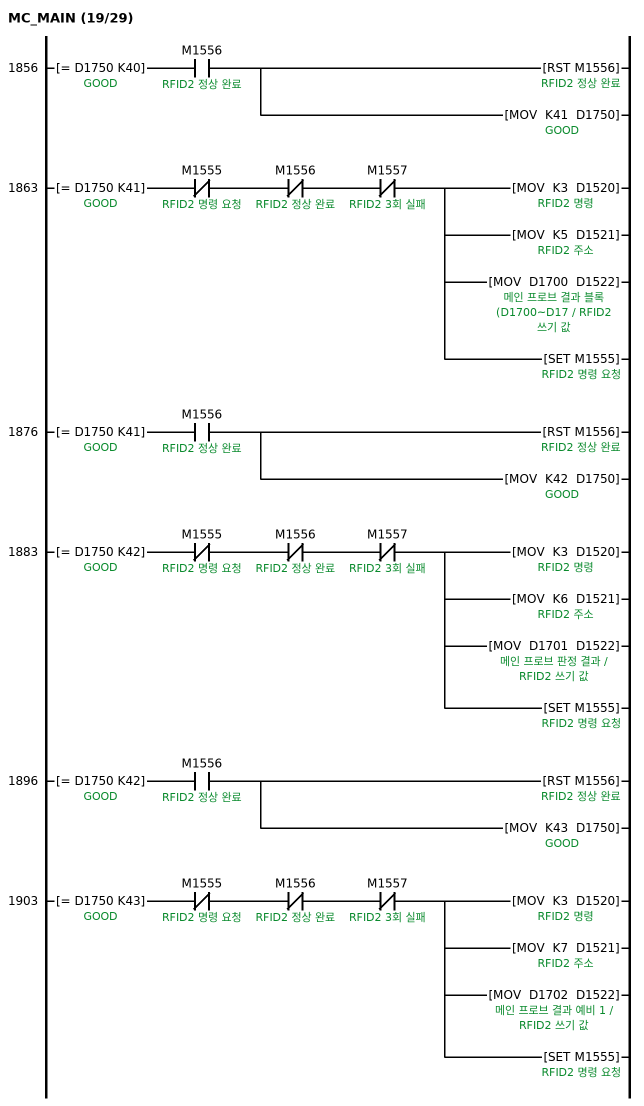
1856  LD=     D1750 K40  ; GOOD
      AND     M1556  ; RFID2 정상 완료
      RST     M1556  ; RFID2 정상 완료
      MOV     K41 D1750
1863  LD=     D1750 K41  ; GOOD
      ANI     M1555  ; RFID2 명령 요청
      ANI     M1556  ; RFID2 정상 완료
      ANI     M1557  ; RFID2 3회 실패
      MOV     K3 D1520
      MOV     K5 D1521
      MOV     D1700 D1522
      SET     M1555  ; RFID2 명령 요청
1876  LD=     D1750 K41  ; GOOD
      AND     M1556  ; RFID2 정상 완료
      RST     M1556  ; RFID2 정상 완료
      MOV     K42 D1750
1883  LD=     D1750 K42  ; GOOD
      ANI     M1555  ; RFID2 명령 요청
      ANI     M1556  ; RFID2 정상 완료
      ANI     M1557  ; RFID2 3회 실패
      MOV     K3 D1520
      MOV     K6 D1521
      MOV     D1701 D1522  ; 메인 프로브 판정 결과
      SET     M1555  ; RFID2 명령 요청
1896  LD=     D1750 K42  ; GOOD
      AND     M1556  ; RFID2 정상 완료
      RST     M1556  ; RFID2 정상 완료
      MOV     K43 D1750
1903  LD=     D1750 K43  ; GOOD
      ANI     M1555  ; RFID2 명령 요청
      ANI     M1556  ; RFID2 정상 완료
      ANI     M1557  ; RFID2 3회 실패
      MOV     K3 D1520
      MOV     K7 D1521
      MOV     D1702 D1522  ; 메인 프로브 결과 예비 1
      SET     M1555  ; RFID2 명령 요청
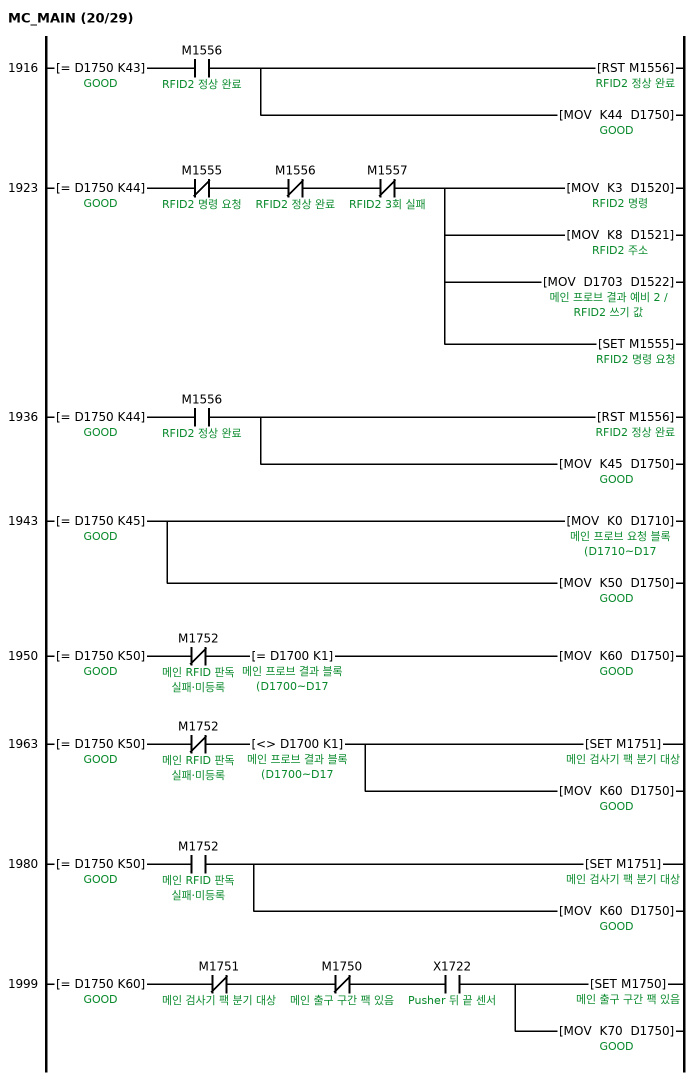
1916  LD=     D1750 K43  ; GOOD
      AND     M1556  ; RFID2 정상 완료
      RST     M1556  ; RFID2 정상 완료
      MOV     K44 D1750
1923  LD=     D1750 K44  ; GOOD
      ANI     M1555  ; RFID2 명령 요청
      ANI     M1556  ; RFID2 정상 완료
      ANI     M1557  ; RFID2 3회 실패
      MOV     K3 D1520
      MOV     K8 D1521
      MOV     D1703 D1522  ; 메인 프로브 결과 예비 2
      SET     M1555  ; RFID2 명령 요청
1936  LD=     D1750 K44  ; GOOD
      AND     M1556  ; RFID2 정상 완료
      RST     M1556  ; RFID2 정상 완료
      MOV     K45 D1750
1943  LD=     D1750 K45  ; GOOD
      MOV     K0 D1710
      MOV     K50 D1750
1950  LD=     D1750 K50  ; GOOD
      ANI     M1752  ; 메인 RFID 판독 실패·미등록
      AND=    D1700 K1  ; 메인 프로브 결과 블록 (D1700~D17
      MOV     K60 D1750
        [note] GOOD
1963  LD=     D1750 K50  ; GOOD
      ANI     M1752  ; 메인 RFID 판독 실패·미등록
      AND<>   D1700 K1  ; 메인 프로브 결과 블록 (D1700~D17
      SET     M1751  ; 메인 검사기 팩 분기 대상
      MOV     K60 D1750
        [note] 2·3·4·5
1980  LD=     D1750 K50  ; GOOD
      AND     M1752  ; 메인 RFID 판독 실패·미등록
      SET     M1751  ; 메인 검사기 팩 분기 대상
      MOV     K60 D1750
        [note] 판독 실패 · 미등록
1999  LD=     D1750 K60  ; GOOD
      ANI     M1751  ; 메인 검사기 팩 분기 대상
      ANI     M1750  ; 메인 출구 구간 팩 있음
      AND     X1722  ; Pusher 뒤 끝 센서
      SET     M1750  ; 메인 출구 구간 팩 있음
      MOV     K70 D1750
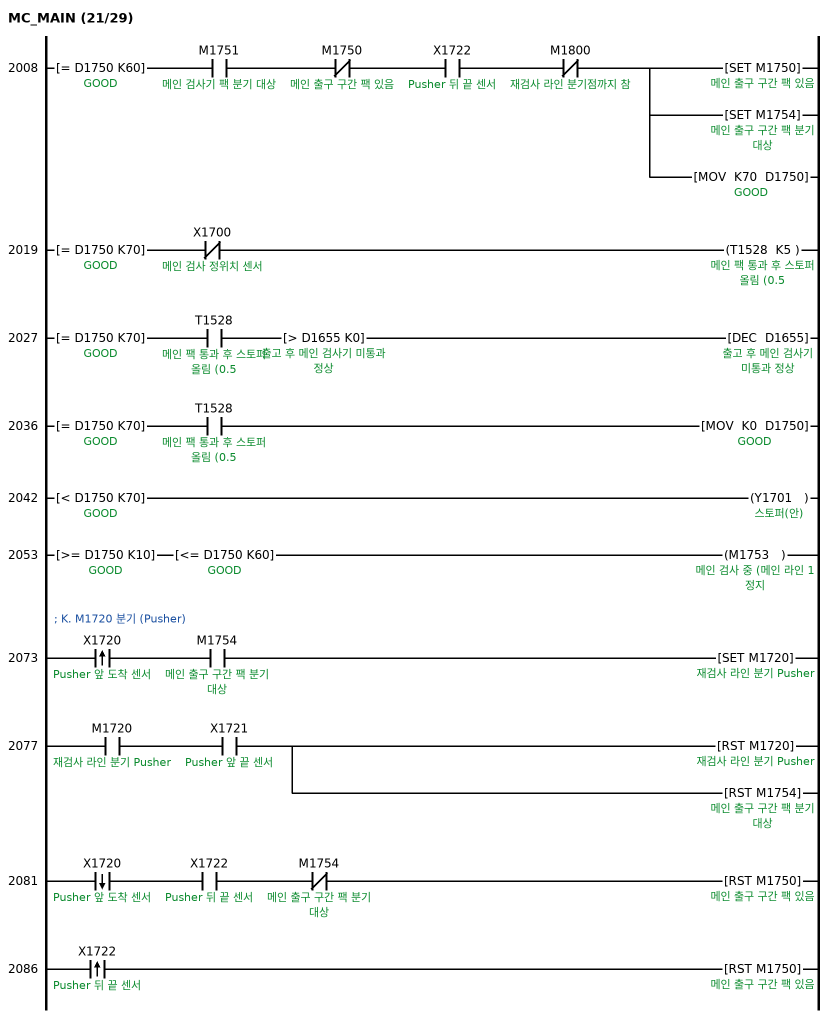
2008  LD=     D1750 K60  ; GOOD
      AND     M1751  ; 메인 검사기 팩 분기 대상
      ANI     M1750  ; 메인 출구 구간 팩 있음
      AND     X1722  ; Pusher 뒤 끝 센서
      ANI     M1800  ; 재검사 라인 분기점까지 참
      SET     M1750  ; 메인 출구 구간 팩 있음
      SET     M1754  ; 메인 출구 구간 팩 분기 대상
      MOV     K70 D1750
2019  LD=     D1750 K70  ; GOOD
      ANI     X1700  ; 메인 검사 정위치 센서
      OUT     T1528 K5  ; 메인 팩 통과 후 스토퍼 올림 (0.5
2027  LD=     D1750 K70  ; GOOD
      AND     T1528  ; 메인 팩 통과 후 스토퍼 올림 (0.5
      AND>    D1655 K0  ; 출고 후 메인 검사기 미통과 정상
      DEC     D1655
2036  LD=     D1750 K70  ; GOOD
      AND     T1528  ; 메인 팩 통과 후 스토퍼 올림 (0.5
      MOV     K0 D1750
2042  LD<     D1750 K70  ; GOOD
      OUT     Y1701  ; 스토퍼(안)
        [note] 스토퍼(안)
2053  LD>=    D1750 K10  ; GOOD
      AND<=   D1750 K60  ; GOOD
      OUT     M1753  ; 메인 검사 중 (메인 라인 1 정지
; K. M1720 분기 (Pusher)
2073  LDP     X1720  ; Pusher 앞 도착 센서
      AND     M1754  ; 메인 출구 구간 팩 분기 대상
      SET     M1720  ; 재검사 라인 분기 Pusher
2077  LD      M1720  ; 재검사 라인 분기 Pusher
      AND     X1721  ; Pusher 앞 끝 센서
      RST     M1720  ; 재검사 라인 분기 Pusher
      RST     M1754  ; 메인 출구 구간 팩 분기 대상
2081  LDF     X1720  ; Pusher 앞 도착 센서
      AND     X1722  ; Pusher 뒤 끝 센서
      ANI     M1754  ; 메인 출구 구간 팩 분기 대상
      RST     M1750  ; 메인 출구 구간 팩 있음
2086  LDP     X1722  ; Pusher 뒤 끝 센서
      RST     M1750  ; 메인 출구 구간 팩 있음
